Staubli VAL3: onStart.pgx

public program onStart(string x_sTrajItem)
  local num l_i
  local num l_nFrameID
  local num l_nToolID
  local num l_nLibNum
  local bool l_bResult
begin
  if sLastTrajItem!=x_sTrajItem
    nPageIndex=0
    nPointIndex=0
  endIf
  call load()
  //
  delay(0)
  sTrajItem=x_sTrajItem
  //

  bBack=false
  for l_i = 0 to size(bBool)-1
    bBool[l_i]=false
  endFor
  //
  for l_i = 0 to size(sList)-1
    sList[l_i]=""
  endFor
  //
  call trajectory:getFrameID(sTrajItem,l_nFrameID)
  call trajectory:getToolID(sTrajItem,l_nToolID)
  call trajectory:getLibName(l_nLibNum,l_bResult)
  call savedata:getFrame(l_nFrameID,fUsingFrame)
  call savedata:getTool(l_nToolID,tUsingTool)
  $jogContext(tUsingTool,fUsingFrame,0)

  sUsingFrame=toString("",l_nFrameID)
  sUsingTool=toString("",l_nToolID)
  sUsingLib=toString("",l_nLibNum)
  logMsg("<traj-jogContext> tool:"+sUsingTool+",frame:"+sUsingFrame)

  sSelPoint=""
  bMark=false



end
